(* IEC 61131-3 sources: PLC-Static-Analysis/modules/plc-rules/src/test/resources/PLCA-L009, 2 files *)

(* ---- compliant.st ---- *)
PROGRAM P_L009ok
VAR
    n : INT;
    m : INT;
    r : REAL;
    b : BOOL;
    c : BOOL;
    q : BOOL;
END_VAR
IF n > 10 THEN
    q := TRUE;
ELSE
    q := FALSE;
END_IF
IF r > 1.0 THEN
    q := TRUE;
ELSIF r < 1.0 THEN
    q := FALSE;
END_IF
END_PROGRAM

(* ---- noncompliant.st ---- *)
PROGRAM P_L009
VAR
    n : INT;
    m : INT;
    r : REAL;
    b : BOOL;
    c : BOOL;
    q : BOOL;
END_VAR
IF n > 10 THEN
    q := TRUE;
ELSIF n <= 10 THEN // PLCA-L009
    q := FALSE;
END_IF
IF n > m THEN
    q := TRUE;
ELSIF m >= n THEN // PLCA-L009
    q := FALSE;
END_IF
END_PROGRAM
